// TIA Portal V21 export
// export: Created 2026-10-12T11:32:16.5280878Z, ExportSetting WithDefaults, DisplayName Totally Integrated Automation Portal, DisplayVersion V21, DisplayName STEP 7 Professional, DisplayVersion V21, DisplayName STEP 7 Safety, DisplayVersion V21, DisplayName Tech WebApplication, DisplayVersion V21, DisplayName WinCC Basic/Comfort/Advanced, DisplayVersion V21, DisplayName WinCC Unified, DisplayVersion V21
DATA_BLOCK "DB_AUTO"   // DB3
{ S7_Optimized_Access := 'FALSE' }
VERSION : 0.1
// stored: AutoNumber true, DBAccessibleFromOPCUA true, IsOnlyStoredInLoadMemory false, IsWriteProtectedInAS false
   VAR
      ACTIVE : Bool;
      "CONVEYOR ON" : Bool;
      "CONVEYOR OFF1" : Bool;
      "CONVEYOR OFF2" : Bool;
      P_TRG : Bool;
      "CAMERA DONE" : Bool;
      "AUTO STATUS" : Int;
      "STOP DELAY TIMER" : IEC_TIMER;
      "SENSOR CHECK DELAY" { S7_SetPoint := 'True'} : IEC_TIMER;
   END_VAR
BEGIN
END_DATA_BLOCK
